TYPE ST_YASKAWA_REF : FB_YASKAWA_REF;
END_TYPE

(* stored: Version 1.1.0.1, ProductVersion 3.1.4024.15
   DUT ST_YASKAWA_REF: Id {175bc9f0-ea60-434c-9653-925d6e7ca1cb} *)
